(* IEC 61131-3 sources: trust-platform/examples/control/03-production-quality-digital-pid/37-discrete-integral-derivative/src, 2 files *)

(* ---- Main.st ---- *)
USING Control;

(* Fraction of the raw-minus-filtered difference applied per update: alpha = dt/(Tf + dt). *)
FUNCTION FilterFraction : LREAL
VAR_INPUT
    CycleTime : LREAL;
    FilterTime : LREAL;
END_VAR
FilterFraction := CycleTime / (FilterTime + CycleTime);
END_FUNCTION

(* One first-order filter update: the filtered value moves alpha of the way toward the raw value. *)
FUNCTION FilterUpdate : LREAL
VAR_INPUT
    PreviousFilteredValue : LREAL;
    RawValue : LREAL;
    FilterFraction : LREAL;
END_VAR
FilterUpdate := PreviousFilteredValue + FilterFraction * (RawValue - PreviousFilteredValue);
END_FUNCTION

FUNCTION SamePidParameters : BOOL
VAR_INPUT
    Left : Control.PIDParameters;
    Right : Control.PIDParameters;
END_VAR
SamePidParameters :=
    Left.ProportionalGain = Right.ProportionalGain
    AND Left.IntegralGain = Right.IntegralGain
    AND Left.DerivativeGain = Right.DerivativeGain
    AND Left.ProportionalSetpointWeight = Right.ProportionalSetpointWeight
    AND Left.DerivativeSetpointWeight = Right.DerivativeSetpointWeight
    AND Left.Bias = Right.Bias
    AND Left.OutputMinimum = Right.OutputMinimum
    AND Left.OutputMaximum = Right.OutputMaximum
    AND Left.RateMinimum = Right.RateMinimum
    AND Left.RateMaximum = Right.RateMaximum
    AND Left.TrackingTime = Right.TrackingTime
    AND Left.AntiWindup = Right.AntiWindup;
END_FUNCTION

PROGRAM Main
VAR
    Controller : Control.PID;
    (* The discrete PID of this lesson: Kp = 16 N·m/rad, Ki = 4 N·m/(rad·s), Kd = 7 N·m·s/rad on the
       filtered angle, the full target change in P, ±20 N·m with back-calculation (Tt = 1 s). *)
    Parameters : Control.PIDParameters := (
        ProportionalGain := LREAL#16.0,
        IntegralGain := LREAL#4.0,
        DerivativeGain := LREAL#7.0,
        ProportionalSetpointWeight := LREAL#1.0,
        DerivativeSetpointWeight := LREAL#0.0,
        Bias := LREAL#0.0,
        OutputMinimum := LREAL#-20.0,
        OutputMaximum := LREAL#20.0,
        RateMinimum := LREAL#-10000.0,
        RateMaximum := LREAL#10000.0,
        TrackingTime := LREAL#1.0,
        AntiWindup := PIDAntiWindup#BackCalculation
    );
    ConfiguredParameters : Control.PIDParameters;
    ParameterRevision : DINT := 0;
    InitialState : Control.PIDInitialState;
    Input : Control.PIDInput;
    Initialized : BOOL := FALSE;
    AutoMode : BOOL := FALSE;
    ManualTorqueNm : LREAL := 0.0;
    SafetyAbort : BOOL := FALSE;
    SetpointRad : LREAL := 0.0;
    AngleRad : LREAL := 0.0;
    VelocityRadS : LREAL := 0.0;
    TorqueNm : LREAL := 0.0;
    (* Drum load of the simulated test rig, in N·m: the loaded trial couples a 2 kg weight at the
       0.1 m drum radius, 1.962 N·m. The controller does not use it. *)
    LoadTorqueNm : LREAL := 0.0;
    (* Measurement filter on the angle: Control.PID differentiates the filtered angle, so D uses the
       filtered velocity. Tf = 0 bypasses the filter; Control Studio applies Tf with the gains. *)
    FilterTimeS : LREAL := 0.1;
    FilterAlpha : LREAL := 1.0;
    FilteredAngleRad : LREAL := 0.0;
    FilterActive : BOOL := FALSE;
    FilterWasActive : BOOL := FALSE;
    (* Project experiment and the positional reading of each controller update (β = 1, γ = 0). *)
    ObservedState : Control.PIDInitialState;
    PreviousFilteredRad : LREAL := 0.0;
    ExperimentEnabled : BOOL := FALSE;
    ExperimentWasEnabled : BOOL := FALSE;
    Active : BOOL := FALSE;
    ErrorRad : LREAL := 0.0;
    ProportionalNm : LREAL := 0.0;
    TrialIntegralNm : LREAL := 0.0;
    DerivativeNm : LREAL := 0.0;
    RequestNm : LREAL := 0.0;
    IntegralNm : LREAL := 0.0;
    (* Software travel and speed limits of the axis. *)
    AngleLimitRad : LREAL := 2.0;
    VelocityLimitRadS : LREAL := 10.0;
    (* Arrival: the measured velocity at the first sample that reaches a new target. *)
    ArrivalSetpointRad : LREAL := 0.0;
    ApproachRad : LREAL := 0.0;
    Arrived : BOOL := TRUE;
    ArrivalVelocityRadS : LREAL := 0.0;
END_VAR

(* Leaving the travel or speed range removes the torque until a full restart. *)
IF ABS(AngleRad) > AngleLimitRad OR ABS(VelocityRadS) > VelocityLimitRadS THEN
    SafetyAbort := TRUE;
END_IF;

(* Control Studio's Apply replaces this complete record at the task boundary. *)
IF NOT Initialized OR NOT SamePidParameters(Left := Parameters, Right := ConfiguredParameters) THEN
    ConfiguredParameters := Parameters;
    ParameterRevision := ParameterRevision + 1;
END_IF;
Controller.Configure(Parameters := Parameters);

IF NOT Initialized THEN
    (* Hot reset: the axis rests without torque and the setpoint follows the measured angle. *)
    ManualTorqueNm := LREAL#0.0;
    IF NOT AutoMode THEN
        SetpointRad := AngleRad;
    END_IF;
    InitialState.Setpoint := SetpointRad;
    InitialState.ProcessValue := AngleRad;
    InitialState.NominalOutput := ManualTorqueNm;
    InitialState.SaturatedOutput := ManualTorqueNm;
    InitialState.SetpointRate := LREAL#0.0;
    InitialState.ProcessValueRate := LREAL#0.0;
    InitialState.FeedForward := LREAL#0.0;
    Controller.Initialize(State := InitialState);
    ArrivalSetpointRad := SetpointRad;
    Initialized := TRUE;
END_IF;

(* Control Studio's project experiment couples the drum load and steps the target to 1.5 rad in Auto.
   Its end uncouples the load and returns to Manual with zero torque. *)
IF ExperimentEnabled AND NOT ExperimentWasEnabled THEN
    Active := TRUE;
    LoadTorqueNm := LREAL#1.962;
    SetpointRad := LREAL#1.5;
    AutoMode := TRUE;
ELSIF NOT ExperimentEnabled AND ExperimentWasEnabled THEN
    Active := FALSE;
    LoadTorqueNm := LREAL#0.0;
    AutoMode := FALSE;
    SetpointRad := AngleRad;
END_IF;
ExperimentWasEnabled := ExperimentEnabled;

(* The filter runs while the controller is in Auto. In Manual and in the Auto-entry scan it restarts
   from the measurement, so entering Auto is exactly bumpless; filtering starts with the next scan. *)
FilterAlpha := FilterFraction(CycleTime := LREAL#0.02, FilterTime := MAX(FilterTimeS, LREAL#0.0));
FilterActive := AutoMode AND NOT SafetyAbort AND Parameters.ProportionalGain > LREAL#0.0;
IF FilterActive AND FilterWasActive THEN
    FilteredAngleRad := FilterUpdate(PreviousFilteredValue := FilteredAngleRad, RawValue := AngleRad, FilterFraction := FilterAlpha);
ELSE
    FilteredAngleRad := AngleRad;
END_IF;
FilterWasActive := FilterActive;

Input.Setpoint := SetpointRad;
Input.ProcessValue := FilteredAngleRad;
Input.CycleTime := LREAL#0.02;
Input.FeedForward := LREAL#0.0;
Input.TrackingOutput := ManualTorqueNm;
IF SafetyAbort THEN
    Input.Mode := PIDMode#Manual;
    Input.ManualOutput := LREAL#0.0;
ELSIF AutoMode AND Parameters.ProportionalGain > LREAL#0.0 THEN
    Input.Mode := PIDMode#Auto;
    Input.ManualOutput := ManualTorqueNm;
ELSE
    Input.Mode := PIDMode#Manual;
    Input.ManualOutput := ManualTorqueNm;
END_IF;
TorqueNm := Controller.Update(Input := Input);

(* The positional reading of this update, in the discrete order: error, P, trial integral, D, request,
   clamp and tracking. Control.PID retains the corrected request; the retained integral is that request
   minus this update's P and D, so the next trial integral starts from it. *)
ObservedState := Controller.GetState();
ErrorRad := SetpointRad - FilteredAngleRad;
ProportionalNm := Parameters.ProportionalGain * ErrorRad;
DerivativeNm := -Parameters.DerivativeGain * (FilteredAngleRad - PreviousFilteredRad) / LREAL#0.02;
TrialIntegralNm := IntegralNm + Parameters.IntegralGain * ErrorRad * LREAL#0.02;
RequestNm := ProportionalNm + TrialIntegralNm + DerivativeNm;
IntegralNm := ObservedState.NominalOutput - ProportionalNm - DerivativeNm;
PreviousFilteredRad := FilteredAngleRad;

IF SetpointRad <> ArrivalSetpointRad THEN
    ArrivalSetpointRad := SetpointRad;
    ApproachRad := SetpointRad - AngleRad;
    Arrived := FALSE;
END_IF;
IF NOT Arrived AND ApproachRad * (SetpointRad - AngleRad) <= LREAL#0.0 THEN
    Arrived := TRUE;
    ArrivalVelocityRadS := VelocityRadS;
END_IF;

END_PROGRAM

CONFIGURATION Config
RESOURCE Res ON PLC
    TASK MainTask(INTERVAL := T#20ms, PRIORITY := 1);
    PROGRAM P1 WITH MainTask : Main;
END_RESOURCE
VAR_CONFIG
    P1.SafetyAbort AT %MX24.0 : BOOL;
    P1.TorqueNm AT %QL0 : LREAL;
    P1.LoadTorqueNm AT %QL8 : LREAL;
    P1.AngleRad AT %IL0 : LREAL;
    P1.VelocityRadS AT %IL8 : LREAL;
    P1.SetpointRad AT %ML0 : LREAL;
    P1.ManualTorqueNm AT %ML8 : LREAL;
    P1.ArrivalVelocityRadS AT %ML16 : LREAL;
    P1.FilteredAngleRad AT %ML32 : LREAL;
    P1.ErrorRad AT %ML40 : LREAL;
    P1.ProportionalNm AT %ML48 : LREAL;
    P1.TrialIntegralNm AT %ML56 : LREAL;
    P1.DerivativeNm AT %ML64 : LREAL;
    P1.RequestNm AT %ML72 : LREAL;
    P1.IntegralNm AT %ML80 : LREAL;
    P1.ExperimentEnabled AT %MX88.0 : BOOL;
    P1.Active AT %MX88.1 : BOOL;
END_VAR
END_CONFIGURATION

(* ---- tests.st ---- *)
(* @trustlsp:runtime-ignore — run these assertions with trust-dev test;
   they are not scheduled PLC instances in the lesson simulator. *)
USING Control;

TEST_PROGRAM TheBenchmarkUpdate
VAR
    ErrorRad : LREAL;
    ProportionalNm : LREAL;
    TrialIntegralNm : LREAL;
    DerivativeNm : LREAL;
    RequestNm : LREAL;
    Controller : Control.PID;
    Parameters : Control.PIDParameters;
    State : Control.PIDInitialState;
    Input : Control.PIDInput;
END_VAR
(* Target 0.50 rad, angle 0.42 rad after 0.40 rad, retained integral 1.962 N·m, Kp 16, Ki 4, Kd 7,
   dt 0.02 s, filter bypassed. *)
ErrorRad := LREAL#0.50 - LREAL#0.42;
ProportionalNm := LREAL#16.0 * ErrorRad;
TrialIntegralNm := LREAL#1.962 + LREAL#4.0 * ErrorRad * LREAL#0.02;
DerivativeNm := LREAL#-7.0 * (LREAL#0.42 - LREAL#0.40) / LREAL#0.02;
RequestNm := ProportionalNm + TrialIntegralNm + DerivativeNm;
ASSERT_NEAR(EXPECTED := LREAL#1.28, ACTUAL := ProportionalNm, DELTA := LREAL#1.0e-12);
ASSERT_NEAR(EXPECTED := LREAL#1.9684, ACTUAL := TrialIntegralNm, DELTA := LREAL#1.0e-12);
ASSERT_NEAR(EXPECTED := LREAL#-7.0, ACTUAL := DerivativeNm, DELTA := LREAL#1.0e-9);
ASSERT_NEAR(EXPECTED := LREAL#-3.7516, ACTUAL := RequestNm, DELTA := LREAL#1.0e-9);
(* Control.PID from the same retained state: the previous update stood at 0.40 rad at rest, so it retained
   P + I + D = 16 · 0.10 + 1.962 + 0 = 3.562 N·m. Its next update gives the same request. *)
Parameters.ProportionalGain := LREAL#16.0;
Parameters.IntegralGain := LREAL#4.0;
Parameters.DerivativeGain := LREAL#7.0;
Parameters.ProportionalSetpointWeight := LREAL#1.0;
Parameters.OutputMinimum := LREAL#-20.0;
Parameters.OutputMaximum := LREAL#20.0;
Parameters.RateMinimum := LREAL#-10000.0;
Parameters.RateMaximum := LREAL#10000.0;
Parameters.TrackingTime := LREAL#1.0;
Parameters.AntiWindup := PIDAntiWindup#BackCalculation;
Controller.Configure(Parameters := Parameters);
State.Setpoint := LREAL#0.50;
State.ProcessValue := LREAL#0.40;
State.NominalOutput := LREAL#3.562;
State.SaturatedOutput := LREAL#3.562;
Controller.Initialize(State := State);
Input.Mode := PIDMode#Auto;
Input.CycleTime := LREAL#0.02;
Input.Setpoint := LREAL#0.50;
Input.ProcessValue := LREAL#0.42;
ASSERT_NEAR(EXPECTED := LREAL#-3.7516, ACTUAL := Controller.Update(Input := Input), DELTA := LREAL#1.0e-9);
END_TEST_PROGRAM

TEST_PROGRAM ClampAndTracking
VAR
    Controller : Control.PID;
    Parameters : Control.PIDParameters;
    State : Control.PIDInitialState;
    Input : Control.PIDInput;
END_VAR
(* A 1.5 rad target step from rest requests P + I* = 16 · 1.5 + 4 · 1.5 · 0.02 = 24.12 N·m: the drive gets
   20 N·m, and tracking corrects the retained request by (dt/Tt)(u_a − u_r) = 0.02 · (20 − 24.12) N·m. *)
Parameters.ProportionalGain := LREAL#16.0;
Parameters.IntegralGain := LREAL#4.0;
Parameters.DerivativeGain := LREAL#7.0;
Parameters.ProportionalSetpointWeight := LREAL#1.0;
Parameters.OutputMinimum := LREAL#-20.0;
Parameters.OutputMaximum := LREAL#20.0;
Parameters.RateMinimum := LREAL#-10000.0;
Parameters.RateMaximum := LREAL#10000.0;
Parameters.TrackingTime := LREAL#1.0;
Parameters.AntiWindup := PIDAntiWindup#BackCalculation;
Controller.Configure(Parameters := Parameters);
Controller.Initialize(State := State);
Input.Mode := PIDMode#Auto;
Input.CycleTime := LREAL#0.02;
Input.Setpoint := LREAL#1.5;
Input.ProcessValue := LREAL#0.0;
ASSERT_NEAR(EXPECTED := LREAL#20.0, ACTUAL := Controller.Update(Input := Input), DELTA := LREAL#1.0e-9);
State := Controller.GetState();
ASSERT_NEAR(EXPECTED := LREAL#24.12 + LREAL#0.02 * (LREAL#20.0 - LREAL#24.12), ACTUAL := State.NominalOutput, DELTA := LREAL#1.0e-9);
END_TEST_PROGRAM
